Fanuc KAREL source: ko00055.KL

-- PROVISIONAL review KL for V770-1; original PC SHA256 0cf5bd195174f7dbd5ea66b0c3fb62ead0bdba51961052277ee288e6b0a9bdf4
-- Incomplete behavior may be omitted. Consult companion uncertainty JSON. Do not deploy.
PROGRAM KO00055
%NOLOCKGROUP
BEGIN
  -- UNRESOLVED_PC offsets 5-12; opcodes 9D,23
  -- UNRESOLVED_PC offsets 17-69; opcodes 27,27,49,7E,AD,27,49,7E,AD,22,31,7E,4A
  -- UNRESOLVED_PC offsets 74-78; opcodes 7F
END KO00055
